// TIA Portal V21 export
FUNCTION_BLOCK "TiaMcpComponentGate"   // FB2, SCL
{ S7_Optimized_Access := 'TRUE' }
VERSION : 0.1
// stored: AutoNumber true, CodeModifiedDate 2026-10-12T06:24:02.9152912Z, CompileDate 2026-10-12T06:24:02.9152912Z, CreationDate 2026-10-12T06:24:10.869627Z, DownloadDate 0001-01-01T00:00:00Z, DownloadWithoutReinit false, HandleErrorsWithinBlock false, ISMultiInstanceCapable true, InterfaceModifiedDate 2026-10-12T06:24:02.4047976Z, IsConsistent true, IsIECCheckEnabled false, IsKnowHowProtected false, IsRetainMemResEnabled false, IsWriteProtected false, LibraryConformanceStatus Das Objekt ist bibliothekskonform., LoadMemoryLength 4307, MemoryReserve 100, ModifiedDate 2026-10-12T06:24:05.9730756Z, PLCSimAdvancedSupport false, ParameterModified 2026-10-12T06:24:02.4047976Z, SetENOAutomatically false, StructureModified 2026-10-12T06:24:02.4047976Z, UDAEnableTagReadback false, VirtualPlcSupport false, WorkMemoryLength 98
   VAR_INPUT
      Enable : Bool;
   END_VAR
   VAR_OUTPUT
      Active : Bool;
   END_VAR
   VAR
      State { S7_SetPoint := 'True'} : "TiaMcpComponentState";
   END_VAR
BEGIN

       #State.Active := #Enable;
       #Active := #State.Active;
END_FUNCTION_BLOCK
